(* IEC 61131-3 sources: Lasal-MCP/examples/SampleSource/LASALScreenAdvancedSolution/LASALScreenAdvancedSolution/LASALScreenAdvacnedSolution/Stations/Terminal/HMI/Class/FileRead, 1 file *)

(* ---- FileRead.st ---- *)
(*!
<Class
	Name               = "FileRead"
	Revision           = "0.0"
	RealtimeTask       = "false"
	CyclicTask         = "false"
	BackgroundTask     = "true"
	DefBackground      = "10 ms"
	Sigmatek           = "false"
	OSInterface        = "false"
	HighPriority       = "false"
	Automatic          = "false"
	UpdateMode         = "Prescan"
	SharedCommandTable = "true"
	Objectsize         = "(444,120)">
	<Channels>
		<Server Name="FileIsCreated" Visualized="false" Initialize="false" WriteProtected="true" Retentive="false"/>
		<Server Name="IntError" Visualized="false" Initialize="false" WriteProtected="true" Retentive="false"/>
		<Server Name="ReadSteps" Visualized="false" Initialize="false" WriteProtected="true" Retentive="false"/>
		<Server Name="StartRead" Visualized="true" Initialize="false" WriteProtected="false" Retentive="false"/>
		<Client Name="_FileSys" Required="false" Internal="false"/>
		<Client Name="_StdLib" Required="false" Internal="false"/>
		<Client Name="StringRAM" Required="true" Internal="false"/>
	</Channels>
</Class>
*)
FileRead : CLASS
	TYPE
	  t_e_ReadSteps :  //! <Type Public="true" Name="t_e_ReadSteps"/>
	  (
	    t_Idle,
	    t_GetFileName,
	    t_Open,
	    t_WaitFileOpen,
	    t_GetLength,
	    t_WaitForGetLength,
	    t_ReadFile,
	    t_WaitForReadFile,
	    t_CloseFile,
	    t_WaitForClose,
	    t_Error
	  )$UDINT;
	END_TYPE
  //Servers:
	ReadSteps 	: SvrChCmd_t_e_ReadSteps_PTofCls_FileRead;
	IntError 	: SvrCh_DINT;
	FileIsCreated 	: SvrCh_DINT;
	StartRead 	: SvrCh_DINT;
  //Clients:
	_FileSys 	: CltChCmd__FileSys;
	_StdLib 	: CltChCmd__StdLib;
	StringRAM 	: CltChCmd_StringRAM;
  //Variables:
		StringLength 	: UDINT;
		FileName : ARRAY [0..99] OF CHAR;

		FunctionID 	: DINT;
		FileHandle 	: DINT;
		FunctionState 	: DINT;
		Length 	: UDINT;
		pReadData 	: ^DINT;
		ReadFile 	: DINT;
		FileIsRead 	: BOOL;
  //Functions:

	FUNCTION VIRTUAL GLOBAL Background
		VAR_INPUT
			EAX 	: UDINT;
		END_VAR
		VAR_OUTPUT
			state (EAX) 	: UDINT;
		END_VAR;

	FUNCTION GLOBAL ReadKoords
		VAR_OUTPUT
			pKoord 	: ^DINT;
		END_VAR;

	FUNCTION GLOBAL GetReadState
		VAR_OUTPUT
			IsRead 	: BOOL;
		END_VAR;

	FUNCTION GLOBAL SetReadState
		VAR_INPUT
			IsDrawing 	: BOOL;
		END_VAR;
  //Tables:
	FUNCTION @STD
		VAR_OUTPUT
			ret_code	: CONFSTATES;
		END_VAR;
	FUNCTION GLOBAL TAB @CT_;
END_CLASS;

#pragma usingLtd _FileSys
#pragma usingLtd _StdLib
#pragma usingLtd StringRAM

FUNCTION VIRTUAL GLOBAL FileRead::Background
	VAR_INPUT
		EAX 	: UDINT;
	END_VAR
	VAR_OUTPUT
		state (EAX) 	: UDINT;
	END_VAR

  //******************************************************************
  //  Read File
  //******************************************************************
  case ReadSteps of

  //******************************************************************
  	t_Idle:

    if (StartRead = 1) then
       StartRead := 0;

       ReadSteps := t_GetFileName;
    end_if;

  //******************************************************************
  	t_GetFileName:

    StringLength := StringRAM.GetLength();

    StringRAM.GetDataAt(pData:= #FileName[0],
                        udSize:= StringLength,
                        udAt:= 0);

    ReadSteps := t_OPEN;

  //******************************************************************
  	t_Open:

    FunctionID := _FileSys.FileOpen_A(Async:= 1,
                                      filename:= #FileName[0],
                                      attributes:= ATT_READ_ONLY);

    ReadSteps := t_WaitFileOpen;

  //*****************************************************************
  	t_WaitFileOpen:

    FunctionState := _FileSys.GetAsyncState(ID:= to_udint(FunctionID),
                                            Erg:= #FileHandle);

      case FunctionState of
        //-----------------------------------
        0:
          if (FileHandle >= 0) then
              ReadSteps := t_GetLength;
          else
            IntError := -1;
            ReadSteps := t_Error;
          end_if;

        //-----------------------------------
        RT_ERG_DELETED,
        RT_INVALID_ID:
          IntError := -2;
          ReadSteps := t_Error;

        //-----------------------------------
        RT_NOT_STARTED,
        RT_IN_PROGRESS:

      end_case;

  //***************************************************************
  	t_GetLength:

    FunctionID := _FileSys.FileLength_A(Async:= 1,
                                        handle:= FileHandle);
    ReadSteps := t_WaitForGetLength;

  //***************************************************************
  	t_WaitForGetLength:

    FunctionState := _FileSys.GetAsyncState(ID:= to_udint(FunctionID),
                                            Erg:= #Length$dint);

    case FunctionState of
      //-----------------------------------
      0:
        if (Length >= 0) then
          ReadSteps := t_ReadFile;
        end_if;

      //-----------------------------------
      RT_ERG_DELETED,
      RT_INVALID_ID:
          IntError := -3;
          ReadSteps := t_Error;

      //-----------------------------------
      RT_NOT_STARTED,
      RT_IN_PROGRESS:

    end_case;

  //**************************************************************
  	t_ReadFile:

    if (pReadData <> NIL) then
      _StdLib.Free(mptr:=pReadData);
    end_if;

    pReadData$^void := _StdLib.Malloc(size:= Length);

    FunctionID$UDINT := _FileSys.FileRead_A(Async:= 1,
                                            handle:= FileHandle,
                                            buffer:= pReadData,
                                            length:= Length);
    ReadSteps := t_WaitForReadFile;

  //**************************************************************
  	t_WaitForReadFile:

    FunctionState := _FileSys.GetAsyncState(ID:= to_udint(FunctionID),
                                            Erg:= #ReadFile);

    case FunctionState of
      //-----------------------------------
      0:
        if (ReadFile >= 0) then
          ReadSteps := t_CloseFile;
        else
          IntError := -4;
          ReadSteps := t_Error;
        end_if;

      //-----------------------------------
      RT_ERG_DELETED,
      RT_INVALID_ID:
        IntError := -5;
        ReadSteps := t_Error;

      //-----------------------------------
      RT_NOT_STARTED,
      RT_IN_PROGRESS:

      end_case;

  //****************************************************************
  	t_CloseFile:

    FunctionID := _FileSys.FileClose_A(Async:= 1,
                                       handle:= FileHandle);

    ReadSteps := t_WaitForClose;

  //****************************************************************
  	t_WaitForClose:

     FunctionState := _FileSys.GetAsyncState(ID:= to_udint(FunctionID),
                                             Erg:= #FileHandle);

     case FunctionState of
        //-----------------------------------
        0:
          if (FileHandle >= 0) then
            FileIsRead := TRUE;
            ReadSteps := t_Idle;
          else
            IntError := -6;
            ReadSteps := t_Error;
          end_if;
     end_case;

  //*****************************************************************
  	t_Error:

  end_case;
  //******************************************************************
  //  End Read File
  //******************************************************************

	state := READY;

END_FUNCTION

FUNCTION GLOBAL FileRead::ReadKoords
	VAR_OUTPUT
		pKoord 	: ^DINT;
	END_VAR

  pKoord := pReadData;

END_FUNCTION

FUNCTION GLOBAL FileRead::GetReadState
	VAR_OUTPUT
		IsRead 	: BOOL;
	END_VAR

  IsRead := FileIsRead;

END_FUNCTION

FUNCTION GLOBAL FileRead::SetReadState
	VAR_INPUT
		IsDrawing 	: BOOL;
	END_VAR

  FileIsRead := IsDrawing;

END_FUNCTION
